(*
SPDX-FileCopyrightText: c 2026 Oleksandr Tiutyk <trofimich@gmail.com>
SPDX-License-Identifier: MIT
License: https://opensource.org/license/mit
*)

(*!
<summary>Checks assigning an empty builder to a populated target without allocating a builder buffer.</summary>
<description>
Uses one task and stays at a stable address while assertions are bound to this instance.
</description>
*)

{attribute 'no_assign'}
{attribute 'no_explicit_call' := 'do not call this function block directly'}
FUNCTION_BLOCK StringBuilderEmptyTest EXTENDS TOF_Testing.SingleCycleTest
VAR_STAT
	{attribute 'hide'}
	_ClassName : STRING := __POUNAME();
END_VAR
VAR
	_Builder : TOF_Core.StringBuilder;
END_VAR

(*!
<summary>Checks assigning an empty builder to a populated target without allocating a builder buffer.</summary>
<description>
The builder is persistent so teardown can release its buffer after an unexpected hook exception.
</description>
*)
METHOD PROTECTED ExecuteTest
VAR
	target : STRING := 'previous contents';
	copied : BOOL;
END_VAR
copied := _Builder.AssignToString(targetString := target);
Assert.ThatBool(
	actual := copied AND_THEN target = '',
	message := "Assigning an empty builder must clear the target and succeed"
).IsTrue();
Assert.ThatBool(
	actual := _Builder.StringLength = 0 AND_THEN _Builder.Capacity = 0,
	message := "Assigning an empty builder must leave it unallocated"
).IsTrue();
END_METHOD

(*!
<summary>Releases the builder buffer before reporting the case result.</summary>
<description>
Safe after partial initialization and after explicit cleanup in the scenario.
</description>
*)
METHOD PROTECTED AfterTest
_Builder.Clear(releaseMemory := TRUE);
END_METHOD

//! <summary>Borrows the concrete class name. Callers must not modify it.</summary>
{attribute 'monitoring' := 'call'}
PROPERTY ClassName : REFERENCE TO STRING
GET
ClassName REF= _ClassName;
END_GET
END_PROPERTY

//! <summary>Borrows the compiler-initialized namespace name. Callers must not modify it.</summary>
{attribute 'monitoring' := 'call'}
PROPERTY NamespaceName : REFERENCE TO STRING
GET
NamespaceName REF= CurrentNamespace.Name;
END_GET
END_PROPERTY

//! <summary>Reports the concrete instance size in bytes.</summary>
{attribute 'monitoring' := 'call'}
PROPERTY SelfSize : ULINT
GET
SelfSize := XSIZEOF(THIS^);
END_GET
END_PROPERTY

END_FUNCTION_BLOCK

(* stored: Version 1.1.0.1
   POU StringBuilderEmptyTest: Id {2ae01f76-1cbd-4d2a-bcae-7c62e3592879}, SpecialFunc None
   Method ExecuteTest: Id {e724b6ab-8cbe-431b-bc74-b7bcc026ce15}
   Method AfterTest: Id {ead87c60-ce3d-4e9f-8a52-cebee0571e52}
   Property ClassName: Id {454184e0-8509-4b7d-8bed-10c5886eb604}
   Get Get: Id {5e0fa7c8-838f-4052-91f0-cd2a21e64321}
   Property NamespaceName: Id {d911d731-19cc-4541-b28e-b4b7ea71aaed}
   Get Get: Id {e7f2ad8c-de43-4a43-917c-72b08a183e6f}
   Property SelfSize: Id {b8ecd9f0-9a63-46fd-9f0f-87712f03ddcb}
   Get Get: Id {40c0a186-2721-4cad-bed1-9e0f419255e6} *)
